(* IEC 61131-3 sources: rusty/tests/lit/correctness, 12 files *)

(* ---- initialization_of_struct_in_function.st ---- *)
// RUN: %COMPILE %s && %RUN | %CHECK %s

TYPE str : STRUCT
    a : DINT := 10; b : DINT := 20; c : DINT := 30; d : DINT;
END_STRUCT END_TYPE

FUNCTION other : DINT
VAR
    a : str;
END_VAR
VAR_INPUT
    index : INT;
END_VAR

    IF index = 0 THEN
        other := a.a;
    ELSIF index = 1 THEN
        other := a.b;
    ELSIF index = 2 THEN
        other := a.c;
    ELSE
        other := a.d;
    END_IF
END_FUNCTION

FUNCTION main : DINT
VAR
    a : DINT;
    b : DINT;
    c : DINT;
    d : DINT;
END_VAR
    a := other(index := 0);
    b := other(index := 1);
    c := other(index := 2);
    d := other(index := 3);

    printf('a=%d$N', a); // CHECK: a=10
    printf('b=%d$N', b); // CHECK: b=20
    printf('c=%d$N', c); // CHECK: c=30
    printf('d=%d$N', d); // CHECK: d=0
END_FUNCTION

(* ---- initialization_of_struct_ref_in_function.st ---- *)
// RUN: %COMPILE %s && %RUN | %CHECK %s

TYPE str : STRUCT
    a : DINT := 10; b : DINT := 20; c : DINT := 30; d : DINT;
END_STRUCT END_TYPE

FUNCTION other : DINT
VAR
    a : str;
END_VAR
VAR_INPUT
    index : INT;
END_VAR

    IF index = 0 THEN
        other := a.a;
    ELSIF index = 1 THEN
        other := a.b;
    ELSIF index = 2 THEN
        other := a.c;
    ELSE
        other := a.d;
    END_IF
END_FUNCTION

FUNCTION main : DINT
VAR
    a : DINT;
    b : DINT;
    c : DINT;
    d : DINT;
END_VAR
    a := other(index := 0);
    b := other(index := 1);
    c := other(index := 2);
    d := other(index := 3);

    printf('a=%d$N', a); // CHECK: a=10
    printf('b=%d$N', b); // CHECK: b=20
    printf('c=%d$N', c); // CHECK: c=30
    printf('d=%d$N', d); // CHECK: d=0
END_FUNCTION

(* ---- boolean_short_circuit.st ---- *)
// RUN: %COMPILE %s && %RUN | %CHECK %s
// Tests that AND_THEN / OR_ELSE short-circuit, and that AND / OR do not.

VAR_GLOBAL
    call_count : DINT;
END_VAR

FUNCTION track : BOOL
VAR_INPUT
    val : BOOL;
END_VAR
    call_count := call_count + 1;
    track := val;
END_FUNCTION

FUNCTION main
    VAR
        result : BOOL;
    END_VAR

    // --- AND_THEN short-circuits when left is FALSE ---
    call_count := 0;
    result := track(FALSE) AND_THEN track(TRUE);
    // CHECK: and_then_false: result=FALSE calls=1
    printf('and_then_false: result=%s calls=%d$N', SEL(result, 'FALSE', 'TRUE'), call_count);

    // --- AND_THEN evaluates right when left is TRUE ---
    call_count := 0;
    result := track(TRUE) AND_THEN track(TRUE);
    // CHECK: and_then_true: result=TRUE calls=2
    printf('and_then_true: result=%s calls=%d$N', SEL(result, 'FALSE', 'TRUE'), call_count);

    // --- AND_THEN returns FALSE when right is FALSE ---
    call_count := 0;
    result := track(TRUE) AND_THEN track(FALSE);
    // CHECK: and_then_right_false: result=FALSE calls=2
    printf('and_then_right_false: result=%s calls=%d$N', SEL(result, 'FALSE', 'TRUE'), call_count);

    // --- OR_ELSE short-circuits when left is TRUE ---
    call_count := 0;
    result := track(TRUE) OR_ELSE track(FALSE);
    // CHECK: or_else_true: result=TRUE calls=1
    printf('or_else_true: result=%s calls=%d$N', SEL(result, 'FALSE', 'TRUE'), call_count);

    // --- OR_ELSE evaluates right when left is FALSE ---
    call_count := 0;
    result := track(FALSE) OR_ELSE track(TRUE);
    // CHECK: or_else_false: result=TRUE calls=2
    printf('or_else_false: result=%s calls=%d$N', SEL(result, 'FALSE', 'TRUE'), call_count);

    // --- OR_ELSE returns FALSE when both are FALSE ---
    call_count := 0;
    result := track(FALSE) OR_ELSE track(FALSE);
    // CHECK: or_else_both_false: result=FALSE calls=2
    printf('or_else_both_false: result=%s calls=%d$N', SEL(result, 'FALSE', 'TRUE'), call_count);

    // --- Contrast: AND evaluates both operands eagerly ---
    call_count := 0;
    result := track(FALSE) AND track(TRUE);
    // CHECK: and_eager: result=FALSE calls=2
    printf('and_eager: result=%s calls=%d$N', SEL(result, 'FALSE', 'TRUE'), call_count);

    // --- Contrast: OR evaluates both operands eagerly ---
    call_count := 0;
    result := track(TRUE) OR track(FALSE);
    // CHECK: or_eager: result=TRUE calls=2
    printf('or_eager: result=%s calls=%d$N', SEL(result, 'FALSE', 'TRUE'), call_count);
END_FUNCTION

(* ---- initialization_of_struct_ref_in_fb_in_function.st ---- *)
// RUN: %COMPILE %s && %RUN | %CHECK %s

TYPE str : STRUCT
    a : DINT := 10; b : DINT := 20; c : DINT := 30; d : DINT;
END_STRUCT END_TYPE

FUNCTION_BLOCK fb
VAR
    a : str;
END_VAR
END_FUNCTION_BLOCK

FUNCTION other : DINT
VAR
    x : fb;
END_VAR
VAR_INPUT
    index : INT;
END_VAR

    IF index = 0 THEN
        other := x.a.a;
    ELSIF index = 1 THEN
        other := x.a.b;
    ELSIF index = 2 THEN
        other := x.a.c;
    ELSE
        other := x.a.d;
    END_IF
END_FUNCTION

FUNCTION main : DINT
VAR
    a : DINT;
    b : DINT;
    c : DINT;
    d : DINT;
END_VAR
    a := other(index := 0);
    b := other(index := 1);
    c := other(index := 2);
    d := other(index := 3);

    printf('a=%d$N', a); // CHECK: a=10
    printf('b=%d$N', b); // CHECK: b=20
    printf('c=%d$N', c); // CHECK: c=30
    printf('d=%d$N', d); // CHECK: d=0
END_FUNCTION

(* ---- array_of_struct_partial_initialization.st ---- *)
// RUN: %COMPILE %s && %RUN | %CHECK %s
// This test verifies that array of struct initialization works correctly
// with different initializer styles:
// 1. Single element initialization in VAR declaration (only first element, rest defaults to zero)
// 2. Full initialization in VAR declaration (all elements explicitly initialized)
// 3. Multiple struct initializers in body assignment

TYPE STRUCT2 :
    STRUCT
        x1 : BOOL;
        x2 : DINT;
        x3 : DINT;
        x4 : DINT;
    END_STRUCT
END_TYPE

PROGRAM mainProg
VAR
    // Single element initializer - only arr1[0] is initialized, arr1[1] should be zeroed
    arr1 : ARRAY[0..1] OF STRUCT2 := [(x1 := TRUE, x2 := 128, x3 := 12, x4 := 421)];
    // Full initializer - both elements explicitly initialized
    arr2 : ARRAY[0..1] OF STRUCT2 := [(x1 := TRUE, x2 := 100), (x1 := FALSE, x2 := 200)];
    // Array for body assignment test
    arr3 : ARRAY[0..1] OF STRUCT2;
END_VAR
    // Multiple struct initializers in body assignment
    arr3 := [(x1 := TRUE, x2 := 500, x3 := 600, x4 := 700), (x1 := FALSE, x2 := 800, x3 := 900, x4 := 1000)];
END_PROGRAM

FUNCTION main : DINT
    mainProg();

    // Check arr1[0] - should have the initialized values
    printf('arr1[0].x1=%d$N', mainProg.arr1[0].x1); // CHECK: arr1[0].x1=1
    printf('arr1[0].x2=%d$N', mainProg.arr1[0].x2); // CHECK: arr1[0].x2=128
    printf('arr1[0].x3=%d$N', mainProg.arr1[0].x3); // CHECK: arr1[0].x3=12
    printf('arr1[0].x4=%d$N', mainProg.arr1[0].x4); // CHECK: arr1[0].x4=421

    // Check arr1[1] - should be zeroed (default initialization)
    printf('arr1[1].x1=%d$N', mainProg.arr1[1].x1); // CHECK: arr1[1].x1=0
    printf('arr1[1].x2=%d$N', mainProg.arr1[1].x2); // CHECK: arr1[1].x2=0
    printf('arr1[1].x3=%d$N', mainProg.arr1[1].x3); // CHECK: arr1[1].x3=0
    printf('arr1[1].x4=%d$N', mainProg.arr1[1].x4); // CHECK: arr1[1].x4=0

    // Check arr2[0] - should have the initialized values, unspecified fields are zero
    printf('arr2[0].x1=%d$N', mainProg.arr2[0].x1); // CHECK: arr2[0].x1=1
    printf('arr2[0].x2=%d$N', mainProg.arr2[0].x2); // CHECK: arr2[0].x2=100
    printf('arr2[0].x3=%d$N', mainProg.arr2[0].x3); // CHECK: arr2[0].x3=0
    printf('arr2[0].x4=%d$N', mainProg.arr2[0].x4); // CHECK: arr2[0].x4=0

    // Check arr2[1] - should have the initialized values, unspecified fields are zero
    printf('arr2[1].x1=%d$N', mainProg.arr2[1].x1); // CHECK: arr2[1].x1=0
    printf('arr2[1].x2=%d$N', mainProg.arr2[1].x2); // CHECK: arr2[1].x2=200
    printf('arr2[1].x3=%d$N', mainProg.arr2[1].x3); // CHECK: arr2[1].x3=0
    printf('arr2[1].x4=%d$N', mainProg.arr2[1].x4); // CHECK: arr2[1].x4=0

    // Check arr3[0] - body assignment with multiple struct initializers
    printf('arr3[0].x1=%d$N', mainProg.arr3[0].x1); // CHECK: arr3[0].x1=1
    printf('arr3[0].x2=%d$N', mainProg.arr3[0].x2); // CHECK: arr3[0].x2=500
    printf('arr3[0].x3=%d$N', mainProg.arr3[0].x3); // CHECK: arr3[0].x3=600
    printf('arr3[0].x4=%d$N', mainProg.arr3[0].x4); // CHECK: arr3[0].x4=700

    // Check arr3[1] - body assignment with multiple struct initializers
    printf('arr3[1].x1=%d$N', mainProg.arr3[1].x1); // CHECK: arr3[1].x1=0
    printf('arr3[1].x2=%d$N', mainProg.arr3[1].x2); // CHECK: arr3[1].x2=800
    printf('arr3[1].x3=%d$N', mainProg.arr3[1].x3); // CHECK: arr3[1].x3=900
    printf('arr3[1].x4=%d$N', mainProg.arr3[1].x4); // CHECK: arr3[1].x4=1000
END_FUNCTION

(* ---- initial_value_in_array_of_struct.st ---- *)
// RUN: %COMPILE %s && %RUN | %CHECK %s

TYPE myStruct : STRUCT
    a, b : DINT;
    c : ARRAY[0..1] OF DINT;
END_STRUCT
END_TYPE

VAR_GLOBAL CONSTANT
    str : myStruct := (a := 50, b := 60, c := [70, 80]);
END_VAR

PROGRAM mainProg
VAR_TEMP
    arr : ARRAY[0..1] OF myStruct := [(a := 10, b := 20, c := [30, 40]), str];
END_VAR
VAR
    a, b, c, d : DINT;
    e, f, g, h : DINT;
END_VAR
    a := arr[0].a;
    b := arr[0].b;
    c := arr[0].c[0];
    d := arr[0].c[1];

    e := arr[1].a;
    f := arr[1].b;
    g := arr[1].c[0];
    h := arr[1].c[1];
END_PROGRAM

FUNCTION main
    mainProg();

    printf('a=%d$N', mainProg.a); // CHECK: a=10
    printf('b=%d$N', mainProg.b); // CHECK: b=20
    printf('c=%d$N', mainProg.c); // CHECK: c=30
    printf('d=%d$N', mainProg.d); // CHECK: d=40
    printf('e=%d$N', mainProg.e); // CHECK: e=50
    printf('f=%d$N', mainProg.f); // CHECK: f=60
    printf('g=%d$N', mainProg.g); // CHECK: g=70
    printf('h=%d$N', mainProg.h); // CHECK: h=80
END_FUNCTION

(* ---- initial_value_in_array_of_struct_body.st ---- *)
// RUN: %COMPILE %s && %RUN | %CHECK %s
// This test verifies that array of struct initialization in the body works correctly
// when the array is declared as VAR_TEMP.
// Case: Full initialization - second element uses a constant struct variable

TYPE myStruct : STRUCT
    a, b : DINT;
    c : ARRAY[0..1] OF DINT;
END_STRUCT
END_TYPE

VAR_GLOBAL CONSTANT
    str : myStruct := (a := 50, b := 60, c := [70, 80]);
END_VAR

PROGRAM mainProg
VAR_TEMP
    arr : ARRAY[0..1] OF myStruct;
END_VAR
VAR
    a, b, c, d : DINT;
    e, f, g, h : DINT;
END_VAR
    arr := [(a := 10, b := 20, c := [30, 40]), str];

    a := arr[0].a;
    b := arr[0].b;
    c := arr[0].c[0];
    d := arr[0].c[1];

    e := arr[1].a;
    f := arr[1].b;
    g := arr[1].c[0];
    h := arr[1].c[1];
END_PROGRAM

FUNCTION main
    mainProg();

    printf('a=%d$N', mainProg.a); // CHECK: a=10
    printf('b=%d$N', mainProg.b); // CHECK: b=20
    printf('c=%d$N', mainProg.c); // CHECK: c=30
    printf('d=%d$N', mainProg.d); // CHECK: d=40
    printf('e=%d$N', mainProg.e); // CHECK: e=50
    printf('f=%d$N', mainProg.f); // CHECK: f=60
    printf('g=%d$N', mainProg.g); // CHECK: g=70
    printf('h=%d$N', mainProg.h); // CHECK: h=80
END_FUNCTION

(* ---- initial_value_in_array_of_struct_body_missing.st ---- *)
// RUN: %COMPILE %s && %RUN | %CHECK %s
// This test verifies that array of struct initialization in the body works correctly
// when the array is declared as VAR_TEMP and only partial elements are provided.
// Case: Missing initialization - only first element is assigned, second should be zero

TYPE myStruct : STRUCT
    a, b : DINT;
    c : ARRAY[0..1] OF DINT;
END_STRUCT
END_TYPE

PROGRAM mainProg
VAR_TEMP
    arr : ARRAY[0..1] OF myStruct;
END_VAR
VAR
    a, b, c, d : DINT;
    e, f, g, h : DINT;
END_VAR
    arr := [(a := 10, b := 20, c := [30, 40])];

    a := arr[0].a;
    b := arr[0].b;
    c := arr[0].c[0];
    d := arr[0].c[1];

    e := arr[1].a;
    f := arr[1].b;
    g := arr[1].c[0];
    h := arr[1].c[1];
END_PROGRAM

FUNCTION main
    mainProg();

    printf('a=%d$N', mainProg.a); // CHECK: a=10
    printf('b=%d$N', mainProg.b); // CHECK: b=20
    printf('c=%d$N', mainProg.c); // CHECK: c=30
    printf('d=%d$N', mainProg.d); // CHECK: d=40
    printf('e=%d$N', mainProg.e); // CHECK: e=0
    printf('f=%d$N', mainProg.f); // CHECK: f=0
    printf('g=%d$N', mainProg.g); // CHECK: g=0
    printf('h=%d$N', mainProg.h); // CHECK: h=0
END_FUNCTION

(* ---- initial_value_in_array_of_struct_body_partial.st ---- *)
// RUN: %COMPILE %s && %RUN | %CHECK %s
// This test verifies that array of struct initialization in the body works correctly
// when the array is declared as VAR_TEMP.
// Case: Partial initialization - second element uses partial struct initializer

TYPE myStruct : STRUCT
    a, b : DINT;
    c : ARRAY[0..1] OF DINT;
END_STRUCT
END_TYPE

PROGRAM mainProg
VAR_TEMP
    arr : ARRAY[0..1] OF myStruct;
END_VAR
VAR
    a, b, c, d : DINT;
    e, f, g, h : DINT;
END_VAR
    arr := [(a := 10, b := 20, c := [30, 40]), (a := 50, c := [70, 80])];

    a := arr[0].a;
    b := arr[0].b;
    c := arr[0].c[0];
    d := arr[0].c[1];

    e := arr[1].a;
    f := arr[1].b;
    g := arr[1].c[0];
    h := arr[1].c[1];
END_PROGRAM

FUNCTION main
    mainProg();

    printf('a=%d$N', mainProg.a); // CHECK: a=10
    printf('b=%d$N', mainProg.b); // CHECK: b=20
    printf('c=%d$N', mainProg.c); // CHECK: c=30
    printf('d=%d$N', mainProg.d); // CHECK: d=40
    printf('e=%d$N', mainProg.e); // CHECK: e=50
    printf('f=%d$N', mainProg.f); // CHECK: f=0
    printf('g=%d$N', mainProg.g); // CHECK: g=70
    printf('h=%d$N', mainProg.h); // CHECK: h=80
END_FUNCTION

(* ---- initial_value_in_array_of_struct_body_var.st ---- *)
// RUN: %COMPILE %s && %RUN | %CHECK %s
// This test verifies that array of struct initialization in the body works correctly.
// This is a companion test to initial_value_in_array_of_struct_body.st which uses VAR_TEMP.
// Case: Full initialization - second element uses a constant struct variable

TYPE myStruct : STRUCT
    a, b : DINT;
    c : ARRAY[0..1] OF DINT;
END_STRUCT
END_TYPE

VAR_GLOBAL CONSTANT
    str : myStruct := (a := 50, b := 60, c := [70, 80]);
END_VAR

PROGRAM mainProg
VAR
    arr : ARRAY[0..1] OF myStruct;
    a, b, c, d : DINT;
    e, f, g, h : DINT;
END_VAR
    arr := [(a := 10, b := 20, c := [30, 40]), str];

    a := arr[0].a;
    b := arr[0].b;
    c := arr[0].c[0];
    d := arr[0].c[1];

    e := arr[1].a;
    f := arr[1].b;
    g := arr[1].c[0];
    h := arr[1].c[1];
END_PROGRAM

FUNCTION main
    mainProg();

    printf('a=%d$N', mainProg.a); // CHECK: a=10
    printf('b=%d$N', mainProg.b); // CHECK: b=20
    printf('c=%d$N', mainProg.c); // CHECK: c=30
    printf('d=%d$N', mainProg.d); // CHECK: d=40
    printf('e=%d$N', mainProg.e); // CHECK: e=50
    printf('f=%d$N', mainProg.f); // CHECK: f=60
    printf('g=%d$N', mainProg.g); // CHECK: g=70
    printf('h=%d$N', mainProg.h); // CHECK: h=80
END_FUNCTION

(* ---- initial_value_in_array_of_struct_body_var_missing.st ---- *)
// RUN: %COMPILE %s && %RUN | %CHECK %s
// This test verifies that array of struct initialization in the body works correctly.
// This is a companion test to initial_value_in_array_of_struct_body_missing.st which uses VAR_TEMP.
// Case: Missing initialization - only first element is assigned, second should be zero

TYPE myStruct : STRUCT
    a, b : DINT;
    c : ARRAY[0..1] OF DINT;
END_STRUCT
END_TYPE

PROGRAM mainProg
VAR
    arr : ARRAY[0..1] OF myStruct;
    a, b, c, d : DINT;
    e, f, g, h : DINT;
END_VAR
    arr := [(a := 10, b := 20, c := [30, 40])];

    a := arr[0].a;
    b := arr[0].b;
    c := arr[0].c[0];
    d := arr[0].c[1];

    e := arr[1].a;
    f := arr[1].b;
    g := arr[1].c[0];
    h := arr[1].c[1];
END_PROGRAM

FUNCTION main
    mainProg();

    printf('a=%d$N', mainProg.a); // CHECK: a=10
    printf('b=%d$N', mainProg.b); // CHECK: b=20
    printf('c=%d$N', mainProg.c); // CHECK: c=30
    printf('d=%d$N', mainProg.d); // CHECK: d=40
    printf('e=%d$N', mainProg.e); // CHECK: e=0
    printf('f=%d$N', mainProg.f); // CHECK: f=0
    printf('g=%d$N', mainProg.g); // CHECK: g=0
    printf('h=%d$N', mainProg.h); // CHECK: h=0
END_FUNCTION

(* ---- initial_value_in_array_of_struct_body_var_partial.st ---- *)
// RUN: %COMPILE %s && %RUN | %CHECK %s
// This test verifies that array of struct initialization in the body works correctly.
// This is a companion test to initial_value_in_array_of_struct_body_partial.st which uses VAR_TEMP.
// Case: Partial initialization - second element uses partial struct initializer

TYPE myStruct : STRUCT
    a, b : DINT;
    c : ARRAY[0..1] OF DINT;
END_STRUCT
END_TYPE

PROGRAM mainProg
VAR
    arr : ARRAY[0..1] OF myStruct;
    a, b, c, d : DINT;
    e, f, g, h : DINT;
END_VAR
    arr := [(a := 10, b := 20, c := [30, 40]), (a := 50, c := [70, 80])];

    a := arr[0].a;
    b := arr[0].b;
    c := arr[0].c[0];
    d := arr[0].c[1];

    e := arr[1].a;
    f := arr[1].b;
    g := arr[1].c[0];
    h := arr[1].c[1];
END_PROGRAM

FUNCTION main
    mainProg();

    printf('a=%d$N', mainProg.a); // CHECK: a=10
    printf('b=%d$N', mainProg.b); // CHECK: b=20
    printf('c=%d$N', mainProg.c); // CHECK: c=30
    printf('d=%d$N', mainProg.d); // CHECK: d=40
    printf('e=%d$N', mainProg.e); // CHECK: e=50
    printf('f=%d$N', mainProg.f); // CHECK: f=0
    printf('g=%d$N', mainProg.g); // CHECK: g=70
    printf('h=%d$N', mainProg.h); // CHECK: h=80
END_FUNCTION
